// TIA Portal V20 export
// export: Created 2026-10-20T18:55:26.6384351Z, ExportSetting None, DisplayName Totally Integrated Automation Portal, DisplayVersion V20 Update 6, DisplayName TIA Portal Openness, DisplayVersion V20 Update 6, DisplayName TIA Portal Version Control Interface, DisplayVersion V20 Update 6, DisplayName SINAMICS Startdrive Advanced, DisplayVersion V20 SP1, DisplayName SINAMICS Startdrive G130, G150, S120, S150, SINAMICS MV, G220, S200, S210, DisplayVersion V20 SP1, DisplayName SINAMICS Startdrive G110M, G120, G120C, G120D, G120P, G115D, DisplayVersion V20 SP1, DisplayName STEP 7 Professional, DisplayVersion V20 Update 6, DisplayName STEP 7 Safety, DisplayVersion V20 Update 2, DisplayName WinCC Basic/Comfort/Advanced, DisplayVersion V20 Update 6, DisplayName WinCC Unified, DisplayVersion V20 Update 6
VAR_GLOBAL   // PLC tag table "IO_Remote_Panel_5"
   "STO VTD - CH1(5)" AT %Q1378.0 : Bool;
   "STO CONVEYOR VTD - CH2(5)" AT %Q1378.3 : Bool;
   "STO CNV VFD (Level 7,8 - Side1) - CH2(5)" AT %Q1384.1 : Bool;
   "STO CNV VFD (Level 1,2,3 - Side1) - CH1(5)" AT %Q1378.4 : Bool;
   "RESET (CABINET)(5)" AT %I1357.3 : Bool;   // Reset (Cabinet) - CH1
   "CABINET COOLING FAN CIRCUIT BREAKER FEEDBACK(5)" AT %I1352.3 : Bool;
   "C5102_SFTY STOPPER ROTATE" AT %Q570.4 : Bool;
   "VTD5 UPPER LIMIT" AT %I1349.0 : Bool;
   "C5103_SFTY STOPPER ROTATE" AT %Q571.0 : Bool;
   "C5106_SFTY STOPPER ROTATE" AT %Q577.4 : Bool;
   "VTD5 SFTY STOPPER CNVS 7,8 - (SIDE 1)" AT %I1371.2 : Bool;
   "STO CNV VFD (Level 4,5,6 - Side1) - CH1(5)" AT %Q1378.6 : Bool;
   "Power Enable Safety Stopper Conveyors (Level 4,5,6 - Side1) - CH1(5)" AT %Q1390.2 : Bool;
   "OVERTRAVEL LOWER LIMIT - CH2(5)" AT %I1357.4 : Bool;   // Overtravel Lower Limit - CH2
   "E-STOP (CABINET) - CH2(5)" AT %I1357.6 : Bool;   // E-Stop (Cabinet) - CH2
   "SCA 5001 STACK LIGHTS YELLOW" AT %Q584.5 : Bool;
   "Chain Slack 1 - CH2(5)" AT %I1364.4 : Bool;   // Chain Slack 1 - CH2
   "CABINET 24V PSU CIRCUIT BREAKER FEEDBACK(5)" AT %I1352.2 : Bool;
   "STO CNV VFD (Level 4,5,6 - Side1) - CH2(5)" AT %Q1378.7 : Bool;
   "C5104 CIRCUIT BREAKER FEEDBACK" AT %I1351.3 : Bool;
   "VTD5 PUSH TO ENTER VTD ZONE" AT %I1350.4 : Bool;
   "Chain Slack 4 - CH1(5)" AT %I1364.3 : Bool;   // Chain Slack 4 - CH1
   "CVTD5 CIRCUIT BREAKER FEEDBACK" AT %I1352.0 : Bool;
   "STO CONVEYOR VTD - CH1(5)" AT %Q1378.2 : Bool;
   "VTD5 CIRCUIT BREAKER FEEDBACK" AT %I1352.1 : Bool;
   "C5103 CIRCUIT BREAKER FEEDBACK" AT %I1351.2 : Bool;
   "Power Enable Safety Stopper Conveyors (Level 7,8 - Side1) - CH2(5)" AT %Q1390.5 : Bool;
   "C5106 CIRCUIT BREAKER FEEDBACK" AT %I1351.5 : Bool;
   "C5105 CIRCUIT BREAKER FEEDBACK" AT %I1351.4 : Bool;
   "C5107_SFTY STOPPER ROTATE" AT %Q578.0 : Bool;
   "C5108_SFTY STOPPER ROTATE" AT %Q578.4 : Bool;
   "STO VTD - CH2(5)" AT %Q1378.1 : Bool;
   "VTD5 LOWER LIMIT" AT %I1349.3 : Bool;
   "VTU HOIST BRAKE SAFETY ENABLE 1(5)" AT %Q1390.6 : Bool;
   "OVERTRAVEL LOWER LIMIT - CH1(5)" AT %I1357.0 : Bool;   // Overtravel Lower Limit - CH1
   "VTD5 SFTY STOPPER CNVS 1,2,3 - (SIDE 1)" AT %I1371.0 : Bool;   // SAFETY STOPPER CONVEYORS (1,2,3 - SIDE 1) EDMFEEDBACK
   "C5102 CIRCUIT BREAKER FEEDBACK" AT %I1351.1 : Bool;
   "VTU HOIST BRAKE SAFETY ENABLE 2(5)" AT %Q1390.7 : Bool;
   "VTD5 PUSH TO EXIT VTD ZONE" AT %I1350.5 : Bool;
   "Power Enable Safety Stopper Conveyors (Level 7,8 - Side1) - CH1(5)" AT %Q1390.4 : Bool;
   "OVERTRAVEL UPPER LIMIT - CH2(5)" AT %I1357.5 : Bool;   // Overtravel Upper Limit - CH2
   "Power Enable Safety Stopper Conveyors (Level 4,5,6 - Side1) - CH2(5)" AT %Q1390.3 : Bool;
   "Chain Slack 2 - CH1(5)" AT %I1364.1 : Bool;   // Chain Slack 2 - CH1
   "Chain Slack 1 - CH1(5)" AT %I1364.0 : Bool;   // Chain Slack 1 - CH1
   "Chain Slack 2 - CH2(5)" AT %I1364.5 : Bool;   // Chain Slack 2 - CH2
   "C5108 CIRCUIT BREAKER FEEDBACK" AT %I1351.7 : Bool;
   "EMERGENCY STOP RESET STATUS - ON(5)" AT %Q585.4 : Bool;   // 920SL1
   "Power Enable Safety Stopper Conveyors (Level 1,2,3 - Side1) - CH2(5)" AT %Q1390.1 : Bool;
   "C5105_SFTY STOPPER ROTATE" AT %Q577.0 : Bool;
   "E-STOP (CABINET) - CH1(5)" AT %I1357.2 : Bool;   // E-Stop (Cabinet)- CH1
   "OVERTRAVEL UPPER LIMIT - CH1(5)" AT %I1357.1 : Bool;   // Overtravel Upper Limit - CH1
   "Chain Slack 3 - CH2(5)" AT %I1364.6 : Bool;   // Chain Slack 3 - CH2
   "C5101_SFTY STOPPER ROTATE" AT %Q570.0 : Bool;
   "STO CNV VFD (Level 1,2,3 - Side1) - CH2(5)" AT %Q1378.5 : Bool;
   "STO CNV VFD (Level 7,8 - Side1) - CH1(5)" AT %Q1384.0 : Bool;
   "C5101 CIRCUIT BREAKER FEEDBACK" AT %I1351.0 : Bool;
   "Chain Slack 4 - CH2(5)" AT %I1364.7 : Bool;   // Chain Slack 4 - CH2
   "C5107 CIRCUIT BREAKER FEEDBACK" AT %I1351.6 : Bool;
   "VTU HOIST BRAKE SAFETY ENABLE EDM FEEDBACK(5)" AT %I1371.3 : Bool;
   "C5104_SFTY STOPPER ROTATE" AT %Q571.4 : Bool;
   "Chain Slack 3 - CH1(5)" AT %I1364.2 : Bool;   // Chain Slack 3 - CH1
   "Power Enable Safety Stopper Conveyors (Level 1,2,3 - Side1) - CH1(5)" AT %Q1390.0 : Bool;
   "VTD5 DOCKING PINS 1 RETRACT" AT %Q585.1 : Bool;
   "VTD5 DOCKING PINS 2 EXTEND" AT %Q585.2 : Bool;
   "SCA 5001 STACK LIGHTS GREEN" AT %Q584.6 : Bool;
   "VTD5 DOCKING PINS 2 RETRACT" AT %Q585.3 : Bool;
   "VTD5 DOCKING PINS 1 EXTEND" AT %Q585.0 : Bool;
   "SCA 5001 STACK LIGHTS RED" AT %Q584.4 : Bool;
   "GATE_SENSOR_CH2(5)" AT %I1371.5 : Bool;
   "VTD5 SFTY STOPPER CNVS 4,5,6 - (SIDE 1)" AT %I1371.4 : Bool;
   "GATE_SENSOR_CH1(5)" AT %I1371.1 : Bool;
END_VAR
